Fanuc KAREL source: kt00110.KL

-- PROVISIONAL review KL for V770-1; original PC SHA256 ecb6cdda3b8208c2fdbc7a852e924b4cad471bec2454f58907e8a7ea11bf4267
-- Incomplete behavior may be omitted. Consult companion uncertainty JSON. Do not deploy.
PROGRAM KT00110
%NOLOCKGROUP
VAR
  R1 : REAL
  OUT : REAL
-- UNRESOLVED_DECL Y2 type=002018
BEGIN
  -- UNRESOLVED_PC offsets 5-16; opcodes 2E,23
  -- UNRESOLVED_PC offsets 21-35; opcodes 2E,22,9D,33,B2
  -- UNRESOLVED_PC offsets 40-63; opcodes 21,22,9D,33,B1,64,6C,23
  -- UNRESOLVED_PC offsets 68-72; opcodes 7F
END KT00110
